// TIA Portal V20 export
Screen "ALARM"  1276x673
  ScreenItem "Button_Back_1" at 2,2 size 90x60  Type=HmiButton
  ScreenItem "Title_ScreenOverview_X390_Y2_1" at 390,2 size 500x30  Type=HmiTextBox
  ScreenItem "Title_ScreenOverview_X390_Y2" at 390,0 size 510x57  Type=HmiTextBox
  ScreenItem "Button_Language" at 97,2 size 90x60  Type=HmiButton
  ScreenItem "permanentareaborderrectangle" at 0,0 size 0x0  Type=HmiRectangle
  ScreenItem "acMessages" at 0,100 size 1276x569  Type=HmiAlarmControl
  ScreenItem "Txt_AlarmClassFilter" at 5,66 size 160x31  Type=HmiSymbolicIOField
  ScreenItem "Btn_AlarmClassFilter" at 167,66 size 109x31  Type=HmiButton
  ScreenItem "Btn_AlarmCodeView" at 1184,2 size 90x60  Type=HmiButton
  ScreenItem "Graphic_BlockedRed" at 1258,5 size 14x14  Type=HmiGraphicView
  ScreenItem "Line_Header_X0_Y64_1" at 0,62 size 1276x0  Type=HmiLine
  ScreenItem "Button_Back" at 2,2 size 90x60  Type=HmiButton
